(* IEC 61131-3 sources: codesys-framework/txt/application/WeVe General (library)/AirPressure/DUT, 1 file *)

(* ---- E_AirPressureState.dut.st ---- *)
{attribute 'qualified_only'}
{attribute 'strict'}
TYPE E_AirPressureState :
(
	OK := 0,
	NOK
);
END_TYPE
